// TIA Portal V21 export
FUNCTION_BLOCK "Batch"   // FB20, GRAPH
TITLE = Batch sequence
// A batch sequence: fill and heat at once, mix, then drain or reject.
   VAR_INPUT
      ACK_EF : Bool;
      start : Bool;
      full : Bool;
      hot : Bool;
      quality : Bool;
      door : Bool;
      overflow : Bool;
      acknowledge : Bool;
      level : Int;
   END_VAR
   VAR_OUTPUT
      valve : Bool;
      lamp : Bool;
      heater : Bool;
      mixer : Bool;
      drain : Bool;
      alarm : Bool;
      clamped : Int;
   END_VAR
BEGIN
// Sequence
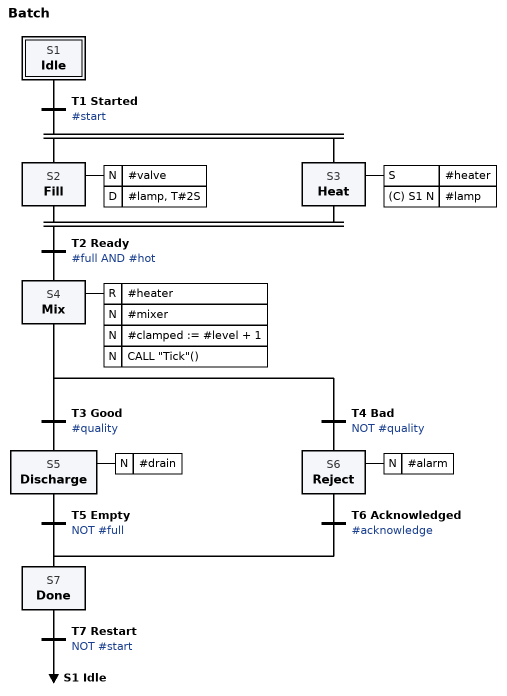
   // permanent pre-instructions
   NETWORK 1
      #lamp := #acknowledge;

   // sequencer 1
   INITIAL_STEP Idle:   // S1
   END_STEP
   TRANSITION Started FROM Idle TO (Fill, Heat)   // T1
      := #start;
   END_TRANSITION
   STEP Fill:   // S2
      supervision V := #overflow;
              N    #valve
              D    #lamp, T#2S
   END_STEP
   STEP Heat:   // S3
      interlock C := #door;
              S    #heater
      (C) S1  N    #lamp
   END_STEP
   TRANSITION Ready FROM (Fill, Heat) TO Mix   // T2
      := #full AND #hot;
   END_TRANSITION
   STEP Mix:   // S4
              R    #heater
              N    #mixer
              N    #clamped := #level + 1
              N    CALL "Tick"()
   END_STEP
   TRANSITION Good FROM Mix TO Discharge   // T3
      := #quality;
   END_TRANSITION
   TRANSITION Bad FROM Mix TO Reject   // T4
      := NOT #quality;
   END_TRANSITION
   STEP Discharge:   // S5
              N    #drain
   END_STEP
   TRANSITION Empty FROM Discharge TO Done   // T5
      := NOT #full;
   END_TRANSITION
   STEP Reject:   // S6
              N    #alarm
   END_STEP
   TRANSITION Acknowledged FROM Reject TO Done   // T6
      := #acknowledge;
   END_TRANSITION
   STEP Done:   // S7
   END_STEP
   TRANSITION Restart FROM Done TO Idle   // T7, jump
      := NOT #start;
   END_TRANSITION

   // permanent post-instructions
   NETWORK 1
      #alarm := #overflow;
END_FUNCTION_BLOCK
